TYPE ST_PolarIIChamber_SelectThreeServiceCtrl :
STRUCT
	Select1 : ST_ServiceCtrl;
	Select2 : ST_ServiceCtrl;
	Select3 : ST_ServiceCtrl;
END_STRUCT
END_TYPE

(* stored: Version 1.1.0.1, ProductVersion 3.1.4026.18
   DUT ST_PolarIIChamber_SelectThreeServiceCtrl: Id {14000000-0000-0000-0000-000000000040} *)
